// TIA Portal V20 export
// export: Created 2026-10-24T18:20:55.1176409Z, ExportSetting WithDefaults, DisplayName Totally Integrated Automation Portal, DisplayVersion V20 Update 6, DisplayName TIA Portal Openness, DisplayVersion V20 Update 6, DisplayName TIA Portal Version Control Interface, DisplayVersion V20 Update 6, DisplayName SINAMICS Startdrive Advanced, DisplayVersion V20 SP1 Update 2, DisplayName SINAMICS Startdrive G110M, G120, G120C, G120D, G120P, G115D, DisplayVersion V20 SP1 Update 2, DisplayName SINAMICS Startdrive G130, G150, S120, S150, SINAMICS MV, G220, S200, S210, DisplayVersion V20 SP1 Update 2, DisplayName STEP 7 Professional, DisplayVersion V20 Update 6, DisplayName STEP 7 Safety, DisplayVersion V20 Update 2, DisplayName WinCC Basic/Comfort/Advanced, DisplayVersion V20 Update 6, DisplayName WinCC Unified, DisplayVersion V20 Update 6
DATA_BLOCK "DB_Machine"   // DB1
TITLE = Machine data
{ S7_Optimized_Access := 'TRUE' }
VERSION : 0.1
// Central data of the filling machine
// stored: AutoNumber true, DBAccessibleFromOPCUA true, DBAccessibleFromWebserver true, IsOnlyStoredInLoadMemory false, IsRetainMemResEnabled false, IsWriteProtectedInAS false, MemoryReserve 100
   VAR
      MachineOn : Bool;   // Machine switched on
      StatusByte : Byte := 16#000F;   // Status bits as byte
      StatusWord : Word := 16#00FF;   // Status bits as word
      StatusDWord : DWord := 16#FFFF;   // Status bits as double word
      StatusLWord : LWord := 16#FFFF_FFFF;   // Status bits as long word
      SmallSigned : SInt := -5;   // Small signed value
      SmallUnsigned : USInt := 200;   // Small unsigned value
      PieceCount : Int;   // Signed piece counter
      PieceCountUnsigned : UInt := 100;   // Unsigned piece counter
      TotalCount : DInt;   // Total number of bottles
      TotalCountUnsigned : UDInt;   // Total number of caps
      LongCount : LInt;   // Long signed counter
      LongCountUnsigned : ULInt;   // Long unsigned counter
      Temperature : Real := 21.5;   // Product temperature in degrees Celsius
      Pressure : LReal := 1.013;   // Line pressure in bar
      CycleTime : Time := T#2S;   // Machine cycle time
      PreciseTime : LTime := LT#500US;   // Precise cycle time
      LegacyTime : S5Time := S5T#10S;   // Legacy time value
      ProductionDate : Date := D#2026-01-01;   // Production date
      ShiftStart : Time_Of_Day := TOD#06:00:00;   // Start of the shift
      PreciseShiftStart : LTime_Of_Day := LTOD#06:00:00.000000001;   // Precise start of the shift
      LegacyTimestamp : Date_And_Time := DT#2026-01-01-06:00:00;   // Legacy time stamp
      PreciseTimestamp : LDT := LDT#2026-01-01-06:00:00;   // Precise time stamp
      Separator : Char := 'A';   // Separator character
      Symbol : WChar := WCHAR#'B';   // Unicode symbol
      MachineName : String[20] := 'Filler';   // Machine name
      OperatorText : WString := WSTRING#'Ready';   // Text for the operator
      LastStart : DTL := DTL#2026-01-01-00:00:00;   // Time of the last start
      Limits : Struct   // Process limits
         Minimum : Real;   // Lower limit
         Maximum : Real := 100.0;   // Upper limit
      END_STRUCT;
      Speeds : Array[0..4] of Int;   // Speed steps
      MainMotor { S7_SetPoint := 'True'} : "UDT_Motor";   // Main drive
      SpeedSetpoint { S7_SetPoint := 'True'} : Real := 50.0;   // Speed setpoint in percent
      InternalState { ExternalAccessible := 'False'; ExternalVisible := 'False'; ExternalWritable := 'False'} : Int;   // Internal state, hidden from HMI and OPC UA
      ReadOnlyValue { ExternalWritable := 'False'} : Real;   // Visible but not writable from HMI and OPC UA
   END_VAR
   VAR RETAIN
      OperatingHours : DInt;   // Operating hours, retentive
      RetainedRecipe : Int := 1;   // Last recipe, retentive
   END_VAR
BEGIN
   Speeds[1] := 10;
   Speeds[2] := 20;
   Speeds[3] := 30;
   Speeds[4] := 40;
END_DATA_BLOCK
